// TIA Portal V21 export
// export: Created 2026-11-22T02:34:34.97806Z, ExportSetting WithDefaults, DisplayName Totally Integrated Automation Portal, DisplayVersion V21 Update 3, DisplayName STEP 7 Professional, DisplayVersion V21 Update 3, DisplayName STEP 7 Safety, DisplayVersion V21, DisplayName Tech WebApplication, DisplayVersion V21, DisplayName WinCC Basic/Comfort/Advanced, DisplayVersion V21 Update 3, DisplayName WinCC Unified, DisplayVersion V21 Update 3
TagTable "C03_Tags"
  D_State : Int  (1 s)
  D_Bool : Bool  (1 s)
  D_SInt : SInt  (1 s)
  D_Int : Int  (1 s)
  D_DInt : DInt  (1 s)
  D_USInt : USInt  (1 s)
  D_UInt : UInt  (1 s)
  D_UDInt : UDInt  (1 s)
  D_Real : Real  (1 s)
  D_LReal : LReal  (1 s)
  D_String : WString  (1 s)
  D_DateTime : DateTime  (1 s)
  D_Pct : Int  (1 s)
  D_Range : Int  (1 s)
  D_Bits : Int  (1 s)
  D_Vis : Bool  (1 s)
  D_En : Bool  (1 s)
  D_X : Int  (1 s)
  D_Y : Int  (1 s)
  D_Max : Real  (1 s)
  D_Min : Real  (1 s)
  D_TL : Int  (1 s)
  D_BarR : Real  (1 s)
